(*
 * Simulacion_Trifasico_MPC_v8_M6_caja_S71200.scl
 *
 * MPC CON LIMITES DE CAMBIO EN TODO EL HORIZONTE ("QP de caja") para S7-1200 (CPU 1212C).
 * Base: el MPC reducido (mismo estimador, mismo termino lineal f, mismos pesos, P = 200, M = 6).
 * En lugar de la solucion sin restricciones + recorte, resuelve en cada ciclo el QP
 *     min 1/2 z'Hz + f'z   con   dumin <= du(k+i) <= dumax  (i = 0..5, las 3 valvulas)
 *                               umin <= u(k) <= umax       (solo el primer movimiento)
 * Todas son cotas de variables ("caja"), y el QP se resuelve con la Hinv que ya usa el MPC:
 * con el conjunto activo A fijo en sus cotas, z = zs + Hinv(:,A) w, con Hinv(A,A) w = cotas - zs(A)
 * (Cholesky de Hinv(A,A)) y multiplicadores = -w. Conjunto activo primal con arranque en caliente
 * (el del ciclo anterior) y TOPE DE 6 ITERACIONES; si se alcanza, el primer movimiento se recorta
 * a sus cotas. Despues, mpc_clipping como en las otras versiones.
 * Frente al MPC completo, deja fuera solo los limites de apertura de los movimientos futuros.
 * Simulacion (escenario de 1000 s): IAE -0.0/+5.1/-0.3 % y variacion total +0.1/+1.3/-0.1 %
 * respecto al MPC completo.
 * [DIAG] mpc_qp_estado: iteraciones usadas (0 = tope); mpc_iter_max; mpc_n_tope.
 * [DIAG] Mediciones de RUNTIME <= 0.0 (vuelta del contador interno) se descartan.
 * LLAMAR DESDE UN OB CICLICO DE 100 ms. Requiere el DB global Diag_HIL.
 *)
DATA_BLOCK PLCGlobalVarMPC
STRUCT
    plc_ts_counter_MPC: DINT;
END_STRUCT
BEGIN
END_DATA_BLOCK
FUNCTION_BLOCK mpc_clipping_MPC
VAR_INPUT
    uk: ARRAY [0..2] OF REAL;
    uk1: ARRAY [0..2] OF REAL;
    b_uoff: ARRAY [0..2] OF REAL;
    b_ny: DINT;
    b_degrees: DINT;
END_VAR
VAR_OUTPUT
    uk_clipped: ARRAY [0..2] OF REAL;
END_VAR
VAR_IN_OUT
    b_Mlim: ARRAY [0..71] OF REAL;   (* solo lectura *)
    b_Mrows: ARRAY [0..71] OF DINT;  (* solo lectura *)
END_VAR
VAR
    nylim: DINT;
    umax: ARRAY [0..2] OF REAL;
    umin: ARRAY [0..2] OF REAL;
    dumin: ARRAY [0..2] OF REAL;
    dumax: ARRAY [0..2] OF REAL;
    iu: DINT;
    du: REAL;
    b_i: DINT;
    tmp: DINT;
    temp1: BOOL;
    temp2: BOOL;
    temp3: BOOL;
END_VAR
nylim := (400 * b_ny) + 1200;
uk_clipped[0] := uk[0];
umax[0] := 3.4028234663852886E+37;
umin[0] := -3.4028234663852886E+37;
dumin[0] := -3.4028234663852886E+37;
dumax[0] := 3.4028234663852886E+37;
uk_clipped[1] := uk[1];
umax[1] := 3.4028234663852886E+37;
umin[1] := -3.4028234663852886E+37;
dumin[1] := -3.4028234663852886E+37;
dumax[1] := 3.4028234663852886E+37;
uk_clipped[2] := uk[2];
umax[2] := 3.4028234663852886E+37;
umin[2] := -3.4028234663852886E+37;
dumin[2] := -3.4028234663852886E+37;
dumax[2] := 3.4028234663852886E+37;
FOR b_i := 0 TO 71 DO
    iu := b_Mrows[b_i];
    temp1 := FALSE;
    temp2 := FALSE;
    temp3 := FALSE;
    IF iu > (nylim - 1200) THEN
        IF iu <= (nylim - 1197) THEN
            iu := (iu - nylim) + 1199;
            umax[iu] := b_Mlim[b_i] + b_uoff[iu];
        ELSE
            temp3 := TRUE;
        END_IF;
    ELSE
        temp3 := TRUE;
    END_IF;
    IF temp3 THEN
        IF iu > (nylim - 600) THEN
            IF iu <= (nylim - 597) THEN
                iu := (iu - nylim) + 599;
                umin[iu] := ( -b_Mlim[b_i]) + b_uoff[iu];
            ELSE
                temp2 := TRUE;
            END_IF;
        ELSE
            temp2 := TRUE;
        END_IF;
    END_IF;
    IF temp2 THEN
        IF iu > nylim THEN
            IF iu <= (nylim + 3) THEN
                dumax[(iu - nylim) - 1] := b_Mlim[b_i];
            ELSE
                temp1 := TRUE;
            END_IF;
        ELSE
            temp1 := TRUE;
        END_IF;
    END_IF;
    IF temp1 THEN
        tmp := nylim + b_degrees;
        IF iu > (tmp - 1) THEN
            IF iu <= (tmp + 2) THEN
                dumin[(iu - nylim) - b_degrees] :=  -b_Mlim[b_i];
            END_IF;
        END_IF;
    END_IF;
END_FOR;
du := uk[0] - uk1[0];
IF du > dumax[0] THEN
    uk_clipped[0] := uk1[0] + dumax[0];
ELSIF du < dumin[0] THEN
    uk_clipped[0] := uk1[0] + dumin[0];
END_IF;
IF uk_clipped[0] > umax[0] THEN
    uk_clipped[0] := umax[0];
ELSIF uk_clipped[0] < umin[0] THEN
    uk_clipped[0] := umin[0];
END_IF;
du := uk[1] - uk1[1];
IF du > dumax[1] THEN
    uk_clipped[1] := uk1[1] + dumax[1];
ELSIF du < dumin[1] THEN
    uk_clipped[1] := uk1[1] + dumin[1];
END_IF;
IF uk_clipped[1] > umax[1] THEN
    uk_clipped[1] := umax[1];
ELSIF uk_clipped[1] < umin[1] THEN
    uk_clipped[1] := umin[1];
END_IF;
du := uk[2] - uk1[2];
IF du > dumax[2] THEN
    uk_clipped[2] := uk1[2] + dumax[2];
ELSIF du < dumin[2] THEN
    uk_clipped[2] := uk1[2] + dumin[2];
END_IF;
IF uk_clipped[2] > umax[2] THEN
    uk_clipped[2] := umax[2];
ELSIF uk_clipped[2] < umin[2] THEN
    uk_clipped[2] := umin[2];
END_IF;
END_FUNCTION_BLOCK
FUNCTION_BLOCK mpcblock_refmd_MPC
VAR_INPUT
    b_ref: ARRAY [0..2] OF REAL;
    b_yoff: ARRAY [0..2] OF REAL;
    b_RYscale: ARRAY [0..2] OF REAL;
END_VAR
VAR_OUTPUT
    rseq: ARRAY [0..2] OF REAL;   (* antes 0..599: solo se usan rseq[0..2] *)
    v: REAL;
END_VAR
VAR
    b_i: DINT;
    ref_0: REAL;
    ref_1: REAL;
    ref_2: REAL;
    b_RYscale_0: REAL;
    b_RYscale_1: REAL;
    b_RYscale_2: REAL;
    b_yoff_0: REAL;
    b_yoff_1: REAL;
    b_yoff_2: REAL;
END_VAR
ref_0 := b_ref[0];
ref_1 := b_ref[1];
ref_2 := b_ref[2];
b_RYscale_0 := b_RYscale[0];
b_RYscale_1 := b_RYscale[1];
b_RYscale_2 := b_RYscale[2];
b_yoff_0 := b_yoff[0];
b_yoff_1 := b_yoff[1];
b_yoff_2 := b_yoff[2];
FOR b_i := 0 TO 0 DO    (* solo rseq[0..2] se usa *)
    rseq[b_i * 3] := (ref_0 * b_RYscale_0) - b_yoff_0;
    rseq[(b_i * 3) + 1] := (ref_1 * b_RYscale_1) - b_yoff_1;
    rseq[(b_i * 3) + 2] := (ref_2 * b_RYscale_2) - b_yoff_2;
END_FOR;
v := 1.0;
END_FUNCTION_BLOCK
FUNCTION_BLOCK MPC_Control
VAR_INPUT
    ssMethodType: INT;
    moorx: ARRAY [0..2] OF REAL;
    b_ref: ARRAY [0..2] OF REAL;
END_VAR
VAR_OUTPUT
    mv: ARRAY [0..2] OF REAL;
END_VAR
VAR
    last_x_PreviousInput: ARRAY [0..6] OF REAL;
    last_mv_DSTATE: ARRAY [0..2] OF REAL;
    c_last_x_InitialCond: ARRAY [0..6] OF REAL := [0.47374550049727165,0.8,0.72,255106.009,0.0,0.0,0.0];
    MPC_3_b_myoff: ARRAY [0..2] OF REAL := [0.8,0.72,3.7];
    MPC_3_b_RYscale: ARRAY [0..2] OF REAL := [1.0,1.0,0.1];
    MPC_3_b_xoff: ARRAY [0..6] OF REAL := [0.47374550049727165,0.8,0.72,255106.009,0.0,0.0,0.0];
    b_a: ARRAY [0..20] OF REAL := [0.0,0.0,0.0,1.0,0.0,0.0,0.0,1.0,0.0,0.0,0.0,1.4503774389728313E-5,0.0,0.0,0.0,0.0,0.0,0.0,0.0,
        0.0,0.0];
    MPC_3_c_a: ARRAY [0..20] OF REAL := [-0.0772292027423523,0.12077646327456022,0.0038948707411090538,1352.9330397447068,
        3.4881337436777948,-1.3447885799979777,-1.1731438171327024,0.269035613232814,0.0038948707411099914,0.09786695730401461,
        348.05070726193321,0.11111867957141662,2.7949959088743932,-2.8155753844244291,0.059593437249509731,0.01962263557286395,
        0.0050480489343075492,14331.413461436903,1.6106730948140586,2.3311020292522353,2.408935193579286];
    MPC_3_b_Mlim: ARRAY [0..71] OF REAL := [0.333871875208127,0.752014397384409,0.515635973890735,0.333871875208127,
        0.752014397384409,0.515635973890735,0.333871875208127,0.752014397384409,0.515635973890735,0.333871875208127,0.752014397384409,
        0.515635973890735,0.333871875208127,0.752014397384409,0.515635973890735,0.333871875208127,0.752014397384409,0.515635973890735,
        0.636128124791873,0.21798560261559102,0.45436402610926496,0.636128124791873,0.21798560261559102,0.45436402610926496,
        0.636128124791873,0.21798560261559102,0.45436402610926496,0.636128124791873,0.21798560261559102,0.45436402610926496,
        0.636128124791873,0.21798560261559102,0.45436402610926496,0.636128124791873,0.21798560261559102,0.45436402610926496,0.035,0.015,
        0.03,0.035,0.015,0.03,0.035,0.015,0.03,0.035,0.015,0.03,0.035,0.015,0.03,0.035,0.015,0.03,0.035,0.015,0.03,0.035,0.015,
        0.03,0.035,0.015,0.03,0.035,0.015,0.03,0.035,0.015,0.03,0.035,0.015,0.03];
    MPC_3_b_Kx: ARRAY [0..125] OF REAL := [-7716.2321024491939,-10901.008671532656,-4264.9443651421188,0.001588040838629834,
        -2543.7442519006345,-1928.3474040587275,19.549174933816971,-44534.108859815329,-44494.776516572136,-26655.405567238093,
        0.0095121063518449449,-8398.6455416316712,-10368.267059564856,158.86185382546796,877.70571831208667,990.07022975809957,
        474.28108255756024,-0.0035701887162486057,96.5496604150103,99.981804413078876,-126.88330315000997,-7621.9188571763643,
        -10775.120625744157,-4206.5654308225376,0.0015700336455973293,-2519.1535379237243,-1907.0052261791157,19.280661326360363,
        -44188.119848216615,-44149.311125111242,-26390.969999054745,0.0094459267062587185,-8342.2703225681144,-10298.597291206755,
        157.85188650166057,864.95022738088733,975.66168439016542,466.81791298662728,-0.0035336819710021609,94.4868041100247,
        97.85316386731445,-125.93879584019494,-7528.1481322542822,-10649.931335099882,-4148.6767278274638,0.0015521046865827432,
        -2494.6400124657093,-1885.7587961853874,19.013959064141872,-43842.116288935795,-43803.826542255309,-26127.843886728973,
        0.0093796925467878947,-8285.8873550992248,-10228.919297363989,156.8419334382582,852.3095979437818,961.384106890396,459.43616436780036,
        -0.003497369852713806,92.447632839384539,95.74911914998566,-124.99418234183436,-7434.9230075303494,-10525.443894660129,
        -4091.2769580451954,0.0015342547665065048,-2470.2045128943837,-1864.6086925692725,18.749068146716176,-43496.122480806749,
        -43458.347088410825,-25866.027371158609,0.0093134067140901722,-8229.4967444644935,-10159.23320514503,155.83198146211291,
        839.78359704931961,947.23718912342133,452.13534732790527,-0.0034612522993006938,90.432068275420264,93.669582511506164,
        -124.04951211934259,-7342.2465048437853,-10401.661341488485,-4034.3648155478659,0.0015164846849855819,-2445.8478788030538,
        -1843.5554965261258,18.485988665509439,-43150.162591337648,-43112.896952629555,-25605.520593125708,0.0092470720701684772,
        -8173.0986508239621,-10089.539209226115,154.82201815145478,827.37198501561852,933.22061617028339,444.91497290855955,
        -0.0034253292477243787,88.440031602080353,91.614465843510473,-123.10483463065196,-7250.1215881048793,-10278.586654731167,
        -3977.9389865477651,0.00149879523623798,-2421.5709518529893,-1822.5997917608677,18.224720801734843,-42804.2606574284,
        -42767.500193326021,-25346.323693295184,0.0091806914982297729,-8116.6932889508143,-10019.83757147498,153.81203184149854,
        815.07451548496078,919.33406638300414,437.7745525706747,-0.0033896006339887937,86.47144350229388,89.5836806634611,
        -122.16019932703135];
    MPC_3_b_Ku1: ARRAY [0..53] OF REAL := [532.9519035819452,1758.7630386838541,-20.218495148255496,1758.7630386838541,
        9920.4082612993716,-164.30092992093171,-20.218495148255496,-164.30092992093171,131.49311423922407,527.80102628666316,
        1737.934860701725,-19.940788232849528,1746.9574860985949,9846.5918503106168,-163.25638356511735,-19.786511752201875,
        -161.71101778484783,130.514941055735,522.666313063715,1717.21838942958,-19.664954679108821,1735.1503109173054,9772.77075083077,
        -162.21185195795246,-19.359488246736596,-159.14605147852319,129.53665804804106,517.54793926655793,1696.6142696551719,
        -19.390994486572826,1723.3415351782228,9698.9487212665517,-161.16732147527,-18.93740822923742,-156.60596908182839,128.55831637410802,
        512.44608071469349,1676.1231380934234,-19.118907749797927,1711.5311924205112,9625.129520129678,-160.12277927000616,
        -18.520255194809877,-154.09070753671722,127.57996718519767,507.36091366067569,1655.7456233405144,-18.848694656201634,
        1699.7193276198914,9551.3169060341625,-159.07821327799945,-18.108012533640888,-151.60020265098143,126.60166162568011];
    MPC_3_b_Kr: ARRAY [0..53] OF REAL := [3186.8373350513389,4275.3677914960599,51.13509990647421,-32.452540397628589,26714.198696645544,72.918687149547608,
        -112.44555961175674,-475.25673471668864,252.72878690712173,3155.2425613858004,4216.8654170260106,50.638144210838703,
        -31.975100691061328,26449.325655557303,72.210143687081711,-110.79080635121332,-467.77820186026861,250.27164490947899,
        3123.8040857581582,4158.8539359264387,50.143499486122451,-31.502311016836352,26185.762042540995,71.504893608304656,
        -109.15217877028672,-460.38123779321489,247.82594499281888,3092.5219240585361,4101.3320539069082,49.651167400702548,
        -31.034149716397167,25923.508020768073,70.802939302930895,-107.52960162200367,-453.06535277614643,245.39169524300604,
        3061.396092190324,4044.2984688129827,49.161149624113243,-30.57059511536292,25662.563753294817,70.104283162373875,
        -105.92299960583885,-445.83005747772961,242.96890375165114,3030.4266060701984,3987.7518705822636,48.673447827046601,
        -30.111625523516803,25402.929403061011,69.408927579747242,-104.33229736767574,-438.67486297920362,240.55757861611488];   (* Kr reducida 18x3 *)
    (* Hinv completa (19 x 19): la usa el QP de caja *)
    MPC_3_b_Hinv: ARRAY [0..360] OF REAL := [0.1702344980572631,-0.000316051953237396,-0.0001214533827540456,-0.036345548841276047,-0.00022994447282000675,
        -7.8535204077971989E-5,-0.035434727013087031,-0.00014382977097906262,-3.4945956300716842E-5,-0.034542309014010772,
        -5.7720706811642746E-5,8.813456011776322E-6,-0.03366968301464044,2.8361008307101794E-5,5.2380161360600679E-5,
        -0.032817675154182616,0.00011438593593406882,9.552481608298865E-5,0.0,-0.000316051953237396,0.010547207252793461,
        2.1132487152157335E-5,-0.0001808791608454948,-0.0023314158969080174,1.0330320315621911E-5,-4.9534035220164727E-5,
        -0.0022413766833578007,1.2191170747377299E-7,7.8036147649309862E-5,-0.0021522792952646508,-9.54953740575078E-6,
        0.00020190252942289518,-0.0020644122541486152,-1.8729858790232883E-5,0.0003221473455128597,-0.0019779594821308214,
        -2.7454115420488076E-5,0.0,-0.0001214533827540456,2.1132487152157335E-5,0.30304411821884769,-6.514990994147179E-5,
        2.1728353827661485E-5,-0.064405415788092474,-8.97885060327611E-6,2.2273463510311548E-5,-0.062989706993492336,
        4.65603793551569E-5,2.2723267969727878E-5,-0.061614542822731315,0.00010110834451599296,2.3046591530932414E-5,
        -0.060282635561179215,0.00015444098334013595,2.322473034505095E-5,-0.058995530723217567,0.0,-0.036345548841276047,
        -0.0001808791608454948,-6.514990994147179E-5,0.17176291685304779,-0.00013612744730930092,-4.4560767159202152E-5,
        -0.0350971665966896,-9.13556293645426E-5,-2.2988766629637194E-5,-0.034463114486899891,-4.65576358502461E-5,
        -9.4991020623304764E-7,-0.033843716347050953,-1.7392388529733022E-6,2.1176229123452892E-5,-0.033239892629933931,
        4.3085064069324768E-5,4.3143636253156359E-5,0.0,-0.00022994447282000675,-0.0023314158969080174,2.1728353827661485E-5,
        -0.00013612744730930092,0.010698246530635966,1.2340538427932472E-5,-4.4760194642908621E-5,-0.0022102015392433554,
        3.4084100679808667E-6,4.4173612422238355E-5,-0.00214976861316072,-5.120830508461208E-6,0.00013070925637258645,
        -0.0020899593246978244,-1.3289405671251868E-5,0.00021489433364024608,-0.0020309671075964997,-2.1128873179308238E-5,
        0.0,-7.8535204077971989E-5,1.0330320315621911E-5,-0.064405415788092474,-4.4560767159202152E-5,1.2340538427932472E-5,
        0.3054148208775625,-1.015071319787011E-5,1.4368446176665112E-5,-0.062417276373171432,2.4179024444158472E-5,
        1.636636500723434E-5,-0.061380921474166857,5.8051555293553663E-5,1.8300251292219083E-5,-0.0603809302382588,
        9.1225498596546247E-5,2.0148793762691288E-5,-0.0594190724227041,0.0,-0.035434727013087031,-4.9534035220164727E-5,
        -8.97885060327611E-6,-0.0350971665966896,-4.4760194642908621E-5,-1.015071319787011E-5,0.17273845134311319,
        -3.9976889795088581E-5,-1.0826124612172019E-5,-0.034391366089294419,-3.5166046909618539E-5,-1.0727884762180431E-5,
        -0.0340234548514619,-3.0316948364924829E-5,-1.0252653775071641E-5,-0.033666135978688227,-2.5428615172775216E-5,
        -9.6634672683266118E-6,0.0,-0.00014382977097906262,-0.0022413766833578007,2.2273463510311548E-5,-9.13556293645426E-5,
        -0.0022102015392433554,1.4368446176665112E-5,-3.9976889795088581E-5,0.010790253977071384,6.7106504165377462E-6,
        1.0310200452023578E-5,-0.002147190141859824,-6.7830888060647946E-7,5.9505058354541645E-5,-0.0021154443640503916,
        -7.8370437343924534E-6,0.00010762063469870516,-0.0020839183592772296,-1.4793606326937087E-5,0.0,
        -3.4945956300716842E-5,1.2191170747377299E-7,-0.062989706993492336,-2.2988766629637194E-5,3.4084100679808667E-6,
        -0.062417276373171432,-1.0826124612172019E-5,6.7106504165377462E-6,0.30702802540700186,1.820897001919164E-6,
        1.005184108764361E-5,-0.061176025329871223,1.4557473121748288E-5,1.3395015801887418E-5,-0.060507679924504308,
        2.7124492071147717E-5,1.6716205009836463E-5,-0.059870813633310996,0.0,-0.034542309014010772,7.8036147649309862E-5,
        4.65603793551569E-5,-0.034463114486899891,4.4173612422238355E-5,2.4179024444158472E-5,-0.034391366089294419,
        1.0310200452023578E-5,1.820897001919164E-6,0.17318140332130527,-2.3547509119607678E-5,-2.0255119613621428E-5,
        -0.03420782335043554,-5.7379181065111574E-5,-4.1654408632959635E-5,-0.034095412692558565,-9.1167816691611789E-5,
        -6.2657366574418234E-5,0.0,-5.7720706811642746E-5,-0.0021522792952646508,2.2723267969727878E-5,-4.65576358502461E-5,
        -0.00214976861316072,1.636636500723434E-5,-3.5166046909618539E-5,-0.002147190141859824,1.005184108764361E-5,
        -2.3547509119607678E-5,0.010824871877124352,3.8016754445631412E-6,-1.1714654534696886E-5,-0.0021406660168113629,
        -2.3487140810286621E-6,3.1080884145891323E-7,-0.0021366194369659398,-8.4238697344242429E-6,0.0,8.813456011776322E-6,
        -9.54953740575078E-6,-0.061614542822731315,-9.4991020623304764E-7,-5.120830508461208E-6,-0.061380921474166857,
        -1.0727884762180431E-5,-6.7830888060647946E-7,-0.061176025329871223,-2.0255119613621428E-5,3.8016754445631412E-6,
        0.30790449828673894,-2.9132918265929341E-5,8.3532488641258142E-6,-0.060660620175687734,-3.7638527243085177E-5,
        1.2949735033266653E-5,-0.060348692971084965,0.0,-0.03366968301464044,0.00020190252942289518,0.00010110834451599296,
        -0.033843716347050953,0.00013070925637258645,5.8051555293553663E-5,-0.0340234548514619,5.9505058354541645E-5,
        1.4557473121748288E-5,-0.03420782335043554,-1.1714654534696886E-5,-2.9132918265929341E-5,0.17311211771562424,
        -8.2943372514784056E-5,-7.26451760390996E-5,-0.034526178406331057,-0.00015415495715396418,-0.00011546864934107219,0.0,
        2.8361008307101794E-5,-0.0020644122541486152,2.3046591530932414E-5,-1.7392388529733022E-6,-0.0020899593246978244,
        1.8300251292219083E-5,-3.0316948364924829E-5,-0.0021154443640503916,1.3395015801887418E-5,-5.7379181065111574E-5,
        -0.0021406660168113629,8.3532488641258142E-6,-8.2943372514784056E-5,0.010803886559746703,3.2103542526533054E-6,
        -0.00010704208143625654,-0.0021887753347569921,-1.9842771425297006E-6,0.0,5.2380161360600679E-5,
        -1.8729858790232883E-5,-0.060282635561179215,2.1176229123452892E-5,-1.3289405671251868E-5,-0.0603809302382588,
        -1.0252653775071641E-5,-7.8370437343924534E-6,-0.060507679924504308,-4.1654408632959635E-5,-2.3487140810286621E-6,
        -0.060660620175687734,-7.26451760390996E-5,3.2103542526533054E-6,0.308065547905881,-0.00010270880655031663,
        8.8847998121922669E-6,-0.0608495071191091,0.0,-0.032817675154182616,0.0003221473455128597,0.00015444098334013595,
        -0.033239892629933931,0.00021489433364024608,9.1225498596546247E-5,-0.033666135978688227,0.00010762063469870516,
        2.7124492071147717E-5,-0.034095412692558565,3.1080884145891323E-7,-3.7638527243085177E-5,-0.034526178406331057,
        -0.00010704208143625654,-0.00010270880655031663,0.17255097784265849,-0.00021442620951791223,-0.00016759605920454502,
        0.0,0.00011438593593406882,-0.0019779594821308214,2.322473034505095E-5,4.3085064069324768E-5,-0.0020309671075964997,
        2.0148793762691288E-5,-2.5428615172775216E-5,-0.0020839183592772296,1.6716205009836463E-5,-9.1167816691611789E-5,
        -0.0021366194369659398,1.2949735033266653E-5,-0.00015415495715396418,-0.0021887753347569921,8.8847998121922669E-6,
        -0.00021442620951791223,0.010729219465504205,4.5706825441767981E-6,0.0,9.552481608298865E-5,-2.7454115420488076E-5,
        -0.058995530723217567,4.3143636253156359E-5,-2.1128873179308238E-5,-0.0594190724227041,-9.6634672683266118E-6,
        -1.4793606326937087E-5,-0.059870813633310996,-6.2657366574418234E-5,-8.4238697344242429E-6,-0.060348692971084965,
        -0.00011546864934107219,-1.9842771425297006E-6,-0.0608495071191091,-0.00016759605920454502,4.5706825441767981E-6,
        0.30753298042695221,0.0,0.0,0.0,0.0,0.0,0.0,0.0,0.0,0.0,0.0,0.0,0.0,0.0,0.0,0.0,0.0,0.0,0.0,0.0,
        9.9999999999999974E-6];
    MPC_3_b_uoff: ARRAY [0..2] OF REAL := [0.656128124791873,0.237985602615591,0.474364026109265];
    MPC_3_b_Mrows: ARRAY [0..71] OF DINT := [1201,1202,1203,1204,1205,1206,1207,1208,1209,1210,1211,1212,1213,1214,1215,1216,1217,
        1218,1801,1802,1803,1804,1805,1806,1807,1808,1809,1810,1811,1812,1813,1814,1815,1816,1817,1818,2401,2402,2403,2404,
        2405,2406,2407,2408,2409,2410,2411,2412,2413,2414,2415,2416,2417,2418,2419,2420,2421,2422,2423,2424,2425,2426,2427,
        2428,2429,2430,2431,2432,2433,2434,2435,2436];
    MPC_3_f_a: ARRAY [0..20] OF REAL := [1.322628327144006E-6,-0.00048116811531683895,-4.3296165052708516E-6,-55.375904267141834,
        0.0,0.0,0.0,-6.9150559684644062E-11,3.7716284508284807E-8,-0.0027971712823564414,-78.996564422017926,0.0,0.0,0.0,
        -2.394037186466665E-10,1.3057639972340998E-7,2.8628831792336135E-7,-273.49234867499621,0.0,0.0,0.0];
    MPC_3_g_a: ARRAY [0..20] OF REAL := [-0.0812759988320282,0.12878974211545094,0.004723574350295019,1608.467976495617,
        3.4881337436777868,-1.3447885799979735,-1.1731438171326984,0.27540380820784305,0.004147779263663315,0.10291146104511424,
        371.46041919189759,0.11111867957141465,2.7949959088743945,-2.8155753844244238,0.065710282048828311,0.023308594370287667,
        0.00655318586773693,16000.578760709672,1.6106730948139927,2.3311020292522739,2.4089351935793255];
    MPC_3_e_a: ARRAY [0..48] OF REAL := [0.9945076508163887,-7.4955911032675407E-6,0.018219343923005435,-0.86686845021470726,0.0,
        0.0,0.0,-0.0054923962532121753,0.99999067551082088,0.018219326989996565,-1.077349693812959,0.0,0.0,0.0,
        -4.0627503649808205E-13,2.2159162199695515E-10,0.99998342284905262,-0.4641225044555104,0.0,0.0,0.0,2.6237854624951297E-12,
        -9.54430195553142E-10,-2.0954813586927272E-9,0.99929334159686478,0.0,0.0,0.0,-6.3159654022047717E-6,0.0022977287773259252,
        2.0675277771461239E-5,264.43732399282771,1.0,0.0,0.0,0.002815004563879495,-1.3684281447907272E-7,2.54613431540441E-5,264.43733847702208,
        0.0,1.0,0.0,2.3147841327022809E-10,-1.26253752403586E-7,-2.7681092818992033E-7,264.43856123334115,0.0,0.0,1.0];
    i0_mpcblock_refmd: mpcblock_refmd_MPC;
    i0_mpc_clipping: mpc_clipping_MPC;
    xk: ARRAY [0..6] OF REAL;
    y_innov: ARRAY [0..2] OF REAL;
    v: REAL;
    rseq: ARRAY [0..2] OF REAL;
    zopt: ARRAY [0..2] OF REAL;
    b_i: DINT;
    rMin: REAL;
    tmp: DINT;
    kDrop: DINT;
    Xnorm0: REAL;
    cMin: REAL;
    cVal: REAL;
    z: ARRAY [0..18] OF REAL;
    t: REAL;
    j_k: DINT;
    rtb_xest: ARRAY [0..6] OF REAL;
    old_u: ARRAY [0..2] OF REAL;
    y_innov_0: REAL;
    D_tmp: DINT;
    (* ---- QP de caja ---- *)
    zs: ARRAY [0..18] OF REAL;        (* solucion sin restricciones -Hinv*f *)
    zq: ARRAY [0..18] OF REAL;        (* solucion del QP de caja *)
    limInf: ARRAY [0..17] OF REAL;    (* cota inferior de cada movimiento *)
    limSup: ARRAY [0..17] OF REAL;    (* cota superior de cada movimiento *)
    actIdx: ARRAY [0..17] OF DINT;    (* conjunto activo: variable fijada *)
    actLado: ARRAY [0..17] OF DINT;   (* -1 en la cota inferior, +1 en la superior *)
    nA: DINT;                         (* tamano del conjunto activo; se conserva entre ciclos *)
    esActiva: ARRAY [0..17] OF BOOL;
    Lch: ARRAY [0..323] OF REAL;      (* factor de Cholesky de Hinv(A,A), 18 x 18 por filas *)
    wv: ARRAY [0..17] OF REAL;
    yv: ARRAY [0..17] OF REAL;
    iterQP: DINT;
    convergio: BOOL;
    peorK: DINT;
    peorV: REAL;
    nuevoI: DINT;
    nuevoLado: DINT;
    sumaQ: REAL;
    ii: DINT;
    jj: DINT;
    kk: DINT;
    pp: DINT;
END_VAR
CASE ssMethodType OF
    0:
        PLCGlobalVarMPC.plc_ts_counter_MPC := 0;
        last_mv_DSTATE[0] := 0.656128124791873;
        last_mv_DSTATE[1] := 0.23798560261559079;
        last_mv_DSTATE[2] := 0.47436402610926476;
        FOR kDrop := 0 TO 6 DO
            last_x_PreviousInput[kDrop] := c_last_x_InitialCond[kDrop];
        END_FOR;
        nA := 0;
    1:
        IF PLCGlobalVarMPC.plc_ts_counter_MPC = 0 THEN
            (* [DIAG] inicio de la medicion *)
            "Diag_HIL".mpc_aux := RUNTIME("Diag_HIL".mpc_mem);

            (* Referencias escaladas *)
            i0_mpcblock_refmd(b_ref := b_ref, b_yoff := MPC_3_b_myoff, b_RYscale := MPC_3_b_RYscale);
            rseq := i0_mpcblock_refmd.rseq;
            v := i0_mpcblock_refmd.v;
            rMin := last_mv_DSTATE[0] - 0.656128124791873;
            Xnorm0 := last_mv_DSTATE[1] - 0.237985602615591;
            cMin := last_mv_DSTATE[2] - 0.474364026109265;

            (* Estimador: innovacion y estado corregido (sin cambios) *)
            FOR kDrop := 0 TO 6 DO
                xk[kDrop] := last_x_PreviousInput[kDrop] - MPC_3_b_xoff[kDrop];
            END_FOR;
            FOR j_k := 0 TO 2 DO
                cVal := 0.0;
                FOR D_tmp := 0 TO 6 DO
                    cVal := (b_a[(3 * D_tmp) + j_k] * xk[D_tmp]) + cVal;
                END_FOR;
                y_innov[j_k] := ((moorx[j_k] * MPC_3_b_RYscale[j_k]) - MPC_3_b_myoff[j_k]) - cVal;
            END_FOR;
            cVal := y_innov[1];
            t := y_innov[0];
            y_innov_0 := y_innov[2];
            FOR j_k := 0 TO 6 DO
                rtb_xest[j_k] := (((MPC_3_c_a[j_k + 7] * cVal) + (MPC_3_c_a[j_k] * t)) + (MPC_3_c_a[j_k + 14] * y_innov_0)
                    ) + xk[j_k];
            END_FOR;

            (* Termino lineal f del QP (z), igual que en el MPC completo *)
            FOR kDrop := 0 TO 18 DO
                z[kDrop] := 0.0;
            END_FOR;
            FOR b_i := 0 TO 17 DO
                cVal := 0.0;
                FOR j_k := 0 TO 6 DO
                    cVal := (MPC_3_b_Kx[(7 * b_i) + j_k] * rtb_xest[j_k]) + cVal;
                END_FOR;
                t := ((MPC_3_b_Kr[3 * b_i] * rseq[0]) + (MPC_3_b_Kr[(3 * b_i) + 1] * rseq[1])) + (MPC_3_b_Kr[(3 * b_i) + 2] * rseq[2]);
                z[b_i] := (((MPC_3_b_Ku1[(3 * b_i) + 1] * Xnorm0) + (MPC_3_b_Ku1[3 * b_i] * rMin)) + (MPC_3_b_Ku1[(3 * b_i)
                     + 2] * cMin)) + (cVal + t);
            END_FOR;

            (* ---------- QP de caja ---------- *)
            (* 1) Solucion sin restricciones zs = -Hinv*f (las 19 variables). Las 3 primeras salen
                  con la misma cuenta que en el MPC reducido. *)
            FOR ii := 0 TO 18 DO
                sumaQ := 0.0;
                FOR jj := 0 TO 18 DO
                    sumaQ := (( -MPC_3_b_Hinv[(19 * jj) + ii]) * z[jj]) + sumaQ;
                END_FOR;
                zs[ii] := sumaQ;
            END_FOR;
            (* 2) Cotas: cambio por muestra en los 6 movimientos de cada valvula y, en el primero,
                  tambien la apertura: umin - u(k-1) <= du(k) <= umax - u(k-1) *)
            FOR ii := 0 TO 17 DO
                limInf[ii] := -MPC_3_b_Mlim[54 + ii];
                limSup[ii] := MPC_3_b_Mlim[36 + ii];
            END_FOR;
            FOR ii := 0 TO 2 DO
                sumaQ := (MPC_3_b_Mlim[ii] + MPC_3_b_uoff[ii]) - last_mv_DSTATE[ii];
                IF sumaQ < limSup[ii] THEN
                    limSup[ii] := sumaQ;
                END_IF;
                sumaQ := ( -MPC_3_b_Mlim[18 + ii] + MPC_3_b_uoff[ii]) - last_mv_DSTATE[ii];
                IF sumaQ > limInf[ii] THEN
                    limInf[ii] := sumaQ;
                END_IF;
            END_FOR;
            (* 3) Conjunto activo: arranca con el del ciclo anterior *)
            FOR ii := 0 TO 17 DO
                esActiva[ii] := FALSE;
            END_FOR;
            FOR kk := 0 TO nA - 1 DO
                esActiva[actIdx[kk]] := TRUE;
            END_FOR;
            FOR ii := 0 TO 18 DO
                zq[ii] := zs[ii];
            END_FOR;
            convergio := FALSE;
            iterQP := 0;
            WHILE (iterQP < 6) AND NOT convergio DO
                iterQP := iterQP + 1;
                (* 3a) w: Hinv(A,A) w = cotas(A) - zs(A), por Cholesky *)
                FOR kk := 0 TO nA - 1 DO
                    IF actLado[kk] < 0 THEN
                        wv[kk] := limInf[actIdx[kk]] - zs[actIdx[kk]];
                    ELSE
                        wv[kk] := limSup[actIdx[kk]] - zs[actIdx[kk]];
                    END_IF;
                END_FOR;
                FOR ii := 0 TO nA - 1 DO
                    FOR jj := 0 TO ii DO
                        sumaQ := MPC_3_b_Hinv[(19 * actIdx[jj]) + actIdx[ii]];
                        FOR pp := 0 TO jj - 1 DO
                            sumaQ := sumaQ - (Lch[(18 * ii) + pp] * Lch[(18 * jj) + pp]);
                        END_FOR;
                        IF ii = jj THEN
                            IF sumaQ <= 1.0E-20 THEN
                                sumaQ := 1.0E-20;
                            END_IF;
                            Lch[(18 * ii) + ii] := SQRT(sumaQ);
                        ELSE
                            Lch[(18 * ii) + jj] := sumaQ / Lch[(18 * jj) + jj];
                        END_IF;
                    END_FOR;
                END_FOR;
                FOR ii := 0 TO nA - 1 DO
                    sumaQ := wv[ii];
                    FOR pp := 0 TO ii - 1 DO
                        sumaQ := sumaQ - (Lch[(18 * ii) + pp] * yv[pp]);
                    END_FOR;
                    yv[ii] := sumaQ / Lch[(18 * ii) + ii];
                END_FOR;
                FOR ii := nA - 1 TO 0 BY -1 DO
                    sumaQ := yv[ii];
                    FOR pp := ii + 1 TO nA - 1 DO
                        sumaQ := sumaQ - (Lch[(18 * pp) + ii] * wv[pp]);
                    END_FOR;
                    wv[ii] := sumaQ / Lch[(18 * ii) + ii];
                END_FOR;
                (* 3b) z = zs + Hinv(:,A) w *)
                FOR ii := 0 TO 18 DO
                    sumaQ := zs[ii];
                    FOR kk := 0 TO nA - 1 DO
                        sumaQ := (MPC_3_b_Hinv[(19 * actIdx[kk]) + ii] * wv[kk]) + sumaQ;
                    END_FOR;
                    zq[ii] := sumaQ;
                END_FOR;
                (* 3c) Multiplicadores (= -w). En la cota inferior deben ser <= 0 y en la superior >= 0:
                       si alguno tiene el signo contrario, se libera el peor *)
                peorK := -1;
                peorV := 1.0E-7;
                FOR kk := 0 TO nA - 1 DO
                    IF actLado[kk] < 0 THEN
                        sumaQ := -wv[kk];
                    ELSE
                        sumaQ := wv[kk];
                    END_IF;
                    IF sumaQ > peorV THEN
                        peorV := sumaQ;
                        peorK := kk;
                    END_IF;
                END_FOR;
                IF peorK >= 0 THEN
                    esActiva[actIdx[peorK]] := FALSE;
                    FOR kk := peorK TO nA - 2 DO
                        actIdx[kk] := actIdx[kk + 1];
                        actLado[kk] := actLado[kk + 1];
                    END_FOR;
                    nA := nA - 1;
                ELSE
                    (* 3d) Variable libre fuera de su cota: se fija la mas violada *)
                    nuevoI := -1;
                    nuevoLado := 0;
                    peorV := 1.0E-7;
                    FOR ii := 0 TO 17 DO
                        IF NOT esActiva[ii] THEN
                            IF (limInf[ii] - zq[ii]) > peorV THEN
                                peorV := limInf[ii] - zq[ii];
                                nuevoI := ii;
                                nuevoLado := -1;
                            ELSIF (zq[ii] - limSup[ii]) > peorV THEN
                                peorV := zq[ii] - limSup[ii];
                                nuevoI := ii;
                                nuevoLado := 1;
                            END_IF;
                        END_IF;
                    END_FOR;
                    IF nuevoI >= 0 THEN
                        actIdx[nA] := nuevoI;
                        actLado[nA] := nuevoLado;
                        esActiva[nuevoI] := TRUE;
                        nA := nA + 1;
                    ELSE
                        convergio := TRUE;
                    END_IF;
                END_IF;
            END_WHILE;
            (* 4) Primer movimiento de cada valvula, dentro de sus cotas (por si se llego al tope) *)
            FOR ii := 0 TO 2 DO
                zopt[ii] := zq[ii];
                IF zopt[ii] > limSup[ii] THEN
                    zopt[ii] := limSup[ii];
                END_IF;
                IF zopt[ii] < limInf[ii] THEN
                    zopt[ii] := limInf[ii];
                END_IF;
            END_FOR;
            IF convergio THEN
                b_i := iterQP;
            ELSE
                b_i := 0;
            END_IF;

            (* [DIAG] estado del QP: iteraciones usadas (0 = se llego al tope de 6) *)
            "Diag_HIL".mpc_qp_estado := b_i;
            "Diag_HIL".mpc_iter_max := MAX(IN1 := "Diag_HIL".mpc_iter_max, IN2 := iterQP);
            IF NOT convergio THEN
                "Diag_HIL".mpc_n_tope := "Diag_HIL".mpc_n_tope + 1;
            END_IF;

            mv[0] := ((last_mv_DSTATE[0] - 0.656128124791873) + zopt[0]) + 0.656128124791873;
            mv[1] := ((last_mv_DSTATE[1] - 0.237985602615591) + zopt[1]) + 0.237985602615591;
            mv[2] := ((last_mv_DSTATE[2] - 0.474364026109265) + zopt[2]) + 0.474364026109265;
            (* Recorte SIEMPRE a los limites del MPC: cambio por muestra (3.5 / 1.5 / 3 %)
               y apertura (2-99 %), con el mismo bloque que usa el MPC completo *)
            old_u[0] := (last_mv_DSTATE[0] - 0.656128124791873) + 0.656128124791873;
            old_u[1] := (last_mv_DSTATE[1] - 0.237985602615591) + 0.237985602615591;
            old_u[2] := (last_mv_DSTATE[2] - 0.474364026109265) + 0.474364026109265;
            i0_mpc_clipping(uk := mv, uk1 := old_u, b_uoff := MPC_3_b_uoff, b_Mlim := MPC_3_b_Mlim, b_Mrows := MPC_3_b_Mrows,
                b_ny := 3, b_degrees := 19);
            mv := i0_mpc_clipping.uk_clipped;

            (* Actualizacion del estimador con la apertura aplicada (sin cambios) *)
            last_mv_DSTATE[0] := mv[0];
            rMin := mv[0] - 0.656128124791873;
            last_mv_DSTATE[1] := mv[1];
            Xnorm0 := mv[1] - 0.237985602615591;
            cMin := mv[2];
            last_mv_DSTATE[2] := mv[2];
            FOR j_k := 0 TO 6 DO
                cVal := 0.0;
                FOR D_tmp := 0 TO 6 DO
                    cVal := (MPC_3_e_a[(7 * D_tmp) + j_k] * xk[D_tmp]) + cVal;
                END_FOR;
                last_x_PreviousInput[j_k] := (((((MPC_3_f_a[j_k + 7] * Xnorm0) + (MPC_3_f_a[j_k] * rMin)) + (MPC_3_f_a[j_k + 14] * (cMin - 0.474364026109265)
                    )) + cVal) + (((MPC_3_g_a[j_k + 7] * y_innov[1]) + (MPC_3_g_a[j_k] * y_innov[0])) + (MPC_3_g_a[j_k + 14] * y_innov[2])
                    )) + MPC_3_b_xoff[j_k];
            END_FOR;

            (* [DIAG] fin de la medicion: tiempo de esta ejecucion en ms *)
            "Diag_HIL".mpc_ms := RUNTIME("Diag_HIL".mpc_mem) * 1000.0;

            (* [DIAG] reinicio de estadisticas desde la tabla de observacion *)
            IF "Diag_HIL".mpc_reset THEN
                "Diag_HIL".mpc_n := 0;
                "Diag_HIL".mpc_sum_ms := 0.0;
                "Diag_HIL".mpc_max_ms := 0.0;
                "Diag_HIL".mpc_iter_max := 0;
                "Diag_HIL".mpc_n_tope := 0;
                "Diag_HIL".mpc_n_infactible := 0;
                "Diag_HIL".mpc_reset := FALSE;
            END_IF;

            (* [DIAG] promedio y maximo desde el ultimo reset *)
            (* [DIAG] Si el contador interno de RUNTIME da la vuelta, la medicion sale <= 0.0 y
               Siemens indica descartarla: solo se acumulan mediciones positivas. *)
            IF "Diag_HIL".mpc_ms > 0.0 THEN
                "Diag_HIL".mpc_n := "Diag_HIL".mpc_n + 1;
                "Diag_HIL".mpc_sum_ms := "Diag_HIL".mpc_sum_ms + "Diag_HIL".mpc_ms;
                "Diag_HIL".mpc_prom_ms := "Diag_HIL".mpc_sum_ms / DINT_TO_LREAL("Diag_HIL".mpc_n);
                "Diag_HIL".mpc_max_ms := MAX(IN1 := "Diag_HIL".mpc_max_ms, IN2 := "Diag_HIL".mpc_ms);
            END_IF;
        END_IF;
        IF PLCGlobalVarMPC.plc_ts_counter_MPC >= 0 THEN   (* divisor desactivado: OB de 100 ms *)
            PLCGlobalVarMPC.plc_ts_counter_MPC := 0;
        ELSE
            PLCGlobalVarMPC.plc_ts_counter_MPC := PLCGlobalVarMPC.plc_ts_counter_MPC + 1;
        END_IF;
END_CASE;
END_FUNCTION_BLOCK
